(* IEC 61131-3 sources: rusty/tests/lit/single/control_statements, 3 files *)

(* ---- if_with_elseif_should_resolve_correctly.st ---- *)
// RUN: %COMPILE %s && %RUN | %CHECK %s
FUNCTION foo : ARRAY[0..1] OF STRING[10]
    VAR
        result : ARRAY[0..1] OF STRING[10];
    END_VAR
    result[0] := 'One';
    result[1] := 'Two';
    foo := result;
END_FUNCTION

FUNCTION getFooResult : STRING[10]
    VAR_INPUT
        index: INT;
    END_VAR
    VAR_IN_OUT
        counterVar : INT;
    END_VAR
    VAR
        fooResult : ARRAY[0..1] OF STRING[10];
    END_VAR
    fooResult := foo();
    counterVar := counterVar + 1;
    getFooResult := fooResult[index];
END_FUNCTION

FUNCTION main
    VAR
        result : INT;
        counterVar: INT;
    END_VAR

    counterVar := 0;

    IF getFooResult(0, counterVar) = 'One' THEN
        result := 1;
    ELSIF getFooResult(1, counterVar) = 'Two' THEN
        result := 2;
    ELSE
        result := 3;
    END_IF

    // CHECK: 1
    printf('%d$N', counterVar);
END_FUNCTION

(* ---- debug_branch_body_locations.st ---- *)
// RUN: %COMPILE_IR %s | %CHECK_IR %s

// A branch body that starts with instructions carrying no location of their own (the
// argument stores of a call) must be attributed to the body's own line, not to the
// location of whatever was generated before it. A body that shares its line with the
// enclosing condition or end keyword gets no line-table row of its own, and a debugger
// cannot then place a breakpoint on it.

FUNCTION_BLOCK Counter
VAR_INPUT step : INT; END_VAR
VAR_OUTPUT total : INT; END_VAR
    total := total + step;
END_FUNCTION_BLOCK

PROGRAM branches
VAR
    c : Counter;
    sel : INT;
    out : INT;
END_VAR
    CASE sel OF
        0: c(step := 1, total => out);
        1: c(step := 2, total => out);
    END_CASE
    IF sel > 0 THEN
        c(step := 3, total => out);
    END_IF
END_PROGRAM

FUNCTION main
    branches();
END_FUNCTION

// Every instruction of a body shares the body's own location, argument stores included.
// CHECK-LABEL: define void @branches
// CHECK: case:
// CHECK: store i16 1, ptr %{{[0-9]+}}, align 2, !dbg ![[CASE0:[0-9]+]]
// CHECK: call void @Counter(ptr %c), !dbg ![[CASE0]]
// CHECK: case1:
// CHECK: store i16 2, ptr %{{[0-9]+}}, align 2, !dbg ![[CASE1:[0-9]+]]
// CHECK: call void @Counter(ptr %c), !dbg ![[CASE1]]
// CHECK: condition_body:
// CHECK: store i16 3, ptr %{{[0-9]+}}, align 2, !dbg ![[IFBODY:[0-9]+]]
// CHECK: call void @Counter(ptr %c), !dbg ![[IFBODY]]

// And that location is the body's source line.
// CHECK-DAG: ![[CASE0]] = !DILocation(line: [[@LINE-25]]
// CHECK-DAG: ![[CASE1]] = !DILocation(line: [[@LINE-25]]
// CHECK-DAG: ![[IFBODY]] = !DILocation(line: [[@LINE-23]]

(* ---- debug_case_body_line_rows.st ---- *)
// REQUIRES: system-linux

// End-to-end: every CASE body keeps a line-table row of its own, which is what lets a
// debugger bind a breakpoint to it. All four bodies here end in the same call and two of
// them are identical, so LLVM's tail merging factors them into shared blocks. A block
// carries one source location, so a merged one is attributed to line 0 and the bodies it
// came from lose their rows.

// RUN: %PLC --debug -Onone -c -o %t.o %s
// RUN: readelf --debug-dump=decodedline %t.o | %CHECK_IR %s

FUNCTION_BLOCK Counter
VAR_INPUT step : INT; reset : BOOL; END_VAR
VAR_OUTPUT total : INT; END_VAR
    IF reset THEN total := 0; ELSE total := total + step; END_IF
END_FUNCTION_BLOCK

PROGRAM branches
VAR
    c : Counter;
    sel : INT;
    out : INT;
END_VAR
    CASE sel OF
        0: c(step := 1, reset := FALSE, total => out); // CHECK-DAG: .st{{ +}}[[@LINE]]{{ +}}
        1: c(step := 2, reset := FALSE, total => out); // CHECK-DAG: .st{{ +}}[[@LINE]]{{ +}}
        2: c(step := 3, reset := TRUE, total => out);  // CHECK-DAG: .st{{ +}}[[@LINE]]{{ +}}
        3: c(step := 1, reset := FALSE, total => out); // CHECK-DAG: .st{{ +}}[[@LINE]]{{ +}}
    END_CASE
END_PROGRAM
